FUNCTION_BLOCK TakeWorkpiece (* Basic Function Block Type *)
  (* Standard: 61499-2 *)
  (* Version 0.0, 7/2/2026, Template *)
  PACKAGE Main;
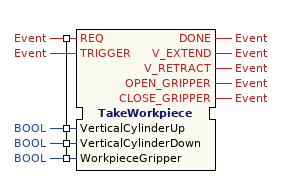
  EVENT_INPUT
    REQ WITH VerticalCylinderUp, VerticalCylinderDown, WorkpieceGripper; (* Normal Execution Request *)
    TRIGGER;
  END_EVENT
  EVENT_OUTPUT
    DONE; (* Initialization Confirm *)
    V_EXTEND; (* Execution Confirmation *)
    V_RETRACT;
    OPEN_GRIPPER;
    CLOSE_GRIPPER;
  END_EVENT
  VAR_INPUT
    VerticalCylinderUp : BOOL; (* Input event qualifier *)
    VerticalCylinderDown : BOOL;
    WorkpieceGripper : BOOL;
  END_VAR
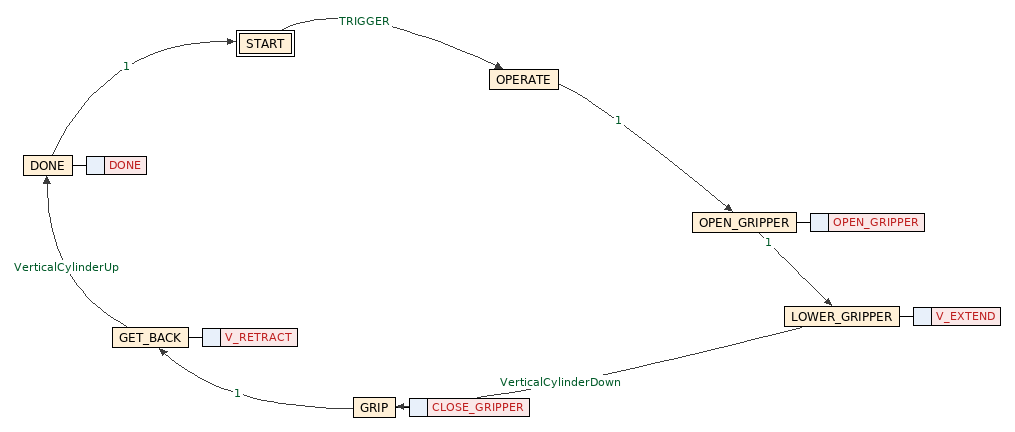
  EC_STATES
    START; (* Initial State *)
    OPERATE;
    OPEN_GRIPPER : -> OPEN_GRIPPER;
    LOWER_GRIPPER : -> V_EXTEND;
    GRIP : -> CLOSE_GRIPPER;
    GET_BACK : -> V_RETRACT;
    DONE : -> DONE;
  END_STATES
  EC_TRANSITIONS
    OPERATE TO OPEN_GRIPPER := 1;
    OPEN_GRIPPER TO LOWER_GRIPPER := 1;
    LOWER_GRIPPER TO GRIP := VerticalCylinderDown;
    GRIP TO GET_BACK := 1;
    GET_BACK TO DONE := VerticalCylinderUp;
    DONE TO START := 1;
    START TO OPERATE := TRIGGER;
  END_TRANSITIONS
  ALGORITHM INIT IN ST: (* Initialization algorithm *)
;
  END_ALGORITHM
  ALGORITHM REQ IN ST: (* Normally executed algorithm *)
;
  END_ALGORITHM
END_FUNCTION_BLOCK
